(*
SPDX-FileCopyrightText: © 2026 Oleksandr Tiutyk <trofimich@gmail.com>
SPDX-License-Identifier: MIT
License: https://opensource.org/license/mit
*)

(*!
<summary>Orders LDATE_AND_TIME values described by generic descriptors.</summary>
<description>
Non-null addresses must reference live LDATE_AND_TIME storage. TypeClass and Size are not validated and no
numeric conversion is performed. Two null addresses compare equal; one null address sorts before a non-null
address. Descriptors are passed by value; payload remains borrowed and is not modified, cloned, released or
retained. IsMemoryOwner does not affect comparison.
</description>
*)

FUNCTION_BLOCK LDateAndTimeComparer EXTENDS TOF_Core.Object IMPLEMENTS TOF_Core.IComparer
VAR_STAT
	//! <summary>Class name shared by all instances of this function block.</summary>
	{attribute 'hide'} 
	_ClassName : STRING := __POUNAME();
END_VAR

{attribute 'monitoring' := 'call'}
PROPERTY ClassName : REFERENCE TO STRING
GET
ClassName REF= _ClassName;
END_GET
END_PROPERTY

(*!
<summary>Compares the first operand with the second using this ordering strategy.</summary>
<description>
Non-null addresses must reference live LDATE_AND_TIME storage. TypeClass and Size are not validated and no
numeric conversion is performed. Two null addresses compare equal; one null address sorts before a non-null
address. Descriptors are passed by value; payload remains borrowed and is not modified, cloned, released or
retained. IsMemoryOwner does not affect comparison. Descendants cannot replace this standard ordering;
implement IComparer separately for a different ordering strategy.
</description>
*)
//!<param name="first">First descriptor; referenced storage is borrowed for the call.</param>
//!<param name="second">Second descriptor; referenced storage is borrowed for the call.</param>
{attribute "object_name" := "Compare"}
METHOD FINAL Compare : TOF_Core.COMPARISON_RESULT
VAR_INPUT
	first : TOF_Core.GENERIC_VALUE;
	second : TOF_Core.GENERIC_VALUE;
END_VAR
VAR
	leftPointer : POINTER TO LDATE_AND_TIME; 
	rightPointer : POINTER TO LDATE_AND_TIME; 
END_VAR
IF first.Address = 0 AND_THEN second.Address = 0 THEN
	Compare := TOF_Core.COMPARISON_RESULT.FIRST_EQUAL_TO_SECOND;
	RETURN;
END_IF

IF first.Address = 0 THEN
	Compare := TOF_Core.COMPARISON_RESULT.FIRST_LESS_THAN_SECOND;
	RETURN;	
END_IF

IF second.Address = 0 THEN
	Compare := TOF_Core.COMPARISON_RESULT.FIRST_GREATER_THAN_SECOND;
	RETURN;	
END_IF

leftPointer := first.Address;
rightPointer := second.Address;

IF leftPointer^ < rightPointer^ THEN
	Compare := TOF_Core.COMPARISON_RESULT.FIRST_LESS_THAN_SECOND;
ELSIF leftPointer^ > rightPointer^ THEN
	Compare := TOF_Core.COMPARISON_RESULT.FIRST_GREATER_THAN_SECOND;
ELSE
	Compare := TOF_Core.COMPARISON_RESULT.FIRST_EQUAL_TO_SECOND;	
END_IF
END_METHOD

{attribute 'monitoring' := 'call'}
PROPERTY NamespaceName : REFERENCE TO STRING
GET
NamespaceName REF= CurrentNamespace.Name;
END_GET
END_PROPERTY

{attribute 'monitoring' := 'call'}
PROPERTY SelfSize : ULINT
GET
SelfSize := XSIZEOF(THIS^);
END_GET
END_PROPERTY

END_FUNCTION_BLOCK

(* stored: Version 1.1.0.1
   POU LDateAndTimeComparer: Id {7fd75ce0-7a6c-46e2-a88f-f44cb5458480}, SpecialFunc None
   Property ClassName: Id {6a172a3e-6ac1-4314-af2e-4424d3c35c1b}
   Get Get: Id {b4eba27d-4bc5-4c2e-b8a0-5d518f0c785f}
   Method Compare: Id {e7e5d810-46d5-4fcb-94f6-62ec678dbe03}
   Property NamespaceName: Id {91e1ec84-f31b-48f5-bc7f-f80fa042348b}
   Get Get: Id {bf4f6d30-1d31-4f2d-b984-bcca3a393db4}
   Property SelfSize: Id {882030fc-f4fd-46cb-a838-4aecc885012e}
   Get Get: Id {27df7169-6dfa-499a-aa6f-6fbe36a27ad8} *)
